(* IEC 61131-3 sources: JingjiangArm/moonboxpro_arm_8.4/Application/Application/任务列表/TensionTask/张力控制/收放料/放料卷径相关/卷径估计, 7 files *)

(* ---- KS_GetFilmThickNessByEstDiaFunc.st ---- *)
(*@CES
Name=KS_GetFilmThickNessByEstDiaFunc
Type=FunctionBlock
TypeGuid=6f9dac99-8de1-4efc-8465-68ac443b7d08
Guid=9700b421-fab0-4030-bfa4-7fb145ef1e2a
HasDeclaration=True
HasImplementation=True
*)
{DECLARATION}
FUNCTION KS_GetFilmThickNessByEstDiaFunc : BOOL
(*2023.12.02.095036 通过估计函数获取料膜厚度@目前主要只应用于接料时的10s不进行卷径补偿部分。
自动获取的方式是
*在开机印刷后超过一定的速度并且处于匀速段
*等待一定的时间后
*持续运行一定的时间后计算这段时间的平均值作为自动的厚度值*)
(*2024.03.16.101611 在停止计算的时候写入初始厚度值|
防止上次料膜太厚计算出的值和本次的薄料厚度差别太大引起异常。厚度值比实际小,对于接料影响会小一些*)
(*2024.7.24.124217 逻辑优化*)
VAR_INPUT
	i_xGetFilmThicknessEn:BOOL;(*自动获取厚度使能@印刷到达一定速度-非调试模式*)
	i_xGetFilmThickNessAuto:BOOL;(*自动获取标志@有效了就通过估计的厚度值获得。无效则通过手动输入获取*)

	i_byWaitTime_Min:BYTE:=1;(*自动满足条件后等待的时间@经过这段时间后开始计算@min*)
	i_byContinuousTime_Min:BYTE:=5;(*持续计算的时间@min*)
	i_byShakeThreshold:BYTE:=10;(*抖动阈值(最值差值法)@丝*)

	i_xEstiThikcknessValid:BOOL;(*估计的厚度值有效*)
	i_rEstiThickness:REAL;(*估计的厚度值@mm*)

	(*2024.03.16.101417*)
	i_rThickness_Init:REAL;(*初始厚度@用于初始化|在退出计算的时候写入该值*)

	i_pxAutoGetDne:POINTER TO BOOL;(*自动获取成功了*)
	i_prThickness:POINTER TO REAL;(*获取的厚度值@mm*)
	i_prTotalThickness:POINTER TO REAL;(*统计的总的厚度值@用于平均处理*)
	i_pudiTotalNum:POINTER TO UDINT;(*统计的次数值@用于平均处理*)
	i_prThickness_Max:POINTER TO REAL;
	i_prThickness_Min:POINTER TO REAL;
	i_ptLastTime:POINTER TO TIME;(*计时使用*)
END_VAR
VAR
	xAutoGetDne: BOOL;
	rThickness: REAL;
	rEstiThickness: REAL;
	rTotalThickness: REAL;
	udiTotalNum: UDINT;
	rThickness_Max: REAL;
	rThickness_Min: REAL;
	rThickness_Manu: REAL;
	tLastTime: TIME;
	tTemp:TIME;
	xEstiThikcknessValid: BOOL;
	rThickness_Init: REAL;(*2024.03.16.101525*)
END_VAR
{IMPLEMENTATION}
(*指针变量写入到临时变量*)
IF i_pxAutoGetDne <>0 THEN
	xAutoGetDne:=i_pxAutoGetDne^;
END_IF
IF i_prThickness<>0 THEN
	rThickness:=i_prThickness^;
END_IF
IF i_prTotalThickness<>0 THEN
	rTotalThickness:=i_prTotalThickness^;
END_IF
IF i_pudiTotalNum<>0 THEN
	udiTotalNum:=i_pudiTotalNum^;
END_IF
IF i_prThickness_Max<>0 THEN
	rThickness_Max:=i_prThickness_Max^;
END_IF
IF i_prThickness_Min<>0 THEN
	rThickness_Min:=i_prThickness_Min^;
END_IF
IF i_ptLastTime<>0 THEN
	tLastTime:=i_ptLastTime^;
END_IF

xEstiThikcknessValid:=i_xEstiThikcknessValid;
rEstiThickness:=i_rEstiThickness;
IF rEstiThickness<=0 OR
	rEstiThickness>=1 THEN(*1MM厚度的几乎没见过，这个只是为了别错的太离谱*)
	xEstiThikcknessValid:=FALSE;(*认为无效|复位所有内容,如果恢复了则重新计算-已经计算完成了就保持吧*)
END_IF

(*2024.03.16.101532*)
rThickness_Init:=i_rThickness_Init;
IF rThickness_Init=0 THEN
	rThickness_Init:=0.02;
END_IF

(*通过估计获取到的厚度值计算*)
(*逻辑处理*)
IF i_xGetFilmThickNessAuto AND(*使用自动获取的方式*)
	xEstiThikcknessValid THEN(*获取估计的厚度值@无效就按照手动输入处理*)
	IF i_xGetFilmThicknessEn AND(*可以自动运算了*)
		NOT xAutoGetDne THEN(*未完成*)
		(*2024.03.16.101150*)
		IF tLastTime=T#0MS THEN(*开始的时候记录时间*)
			tLastTime:=TIME();
		END_IF

		tTemp:=DWORD_TO_TIME(BYTE_TO_DWORD(i_byWaitTime_Min)*60*1000);(*转换为ms*)
		IF TIME()-tLastTime>tTemp THEN(*等待时间够了*)
			tTemp:=DWORD_TO_TIME(BYTE_TO_DWORD(i_byWaitTime_Min+i_byContinuousTime_Min)*60*1000);(*转换为ms*)
			(*累计厚度值*)
			udiTotalNum:=udiTotalNum+1;
			rTotalThickness:=rTotalThickness+rEstiThickness;
			(*记录最大值和最小值*)
			IF rThickness_Max<rEstiThickness THEN
				rThickness_Max:=rEstiThickness;
			END_IF
			IF rThickness_Min>rEstiThickness THEN
				rThickness_Min:=rEstiThickness;
			END_IF

			(*记录的时间到了@检查最大和最小值偏差是否符合要求*)
			IF TIME()-tLastTime>tTemp THEN
				(*符和要求|写入*)
				IF (rThickness_Max-rThickness_Min)<=BYTE_TO_REAL(i_byShakeThreshold)/100.0 THEN
					IF udiTotalNum<>0 THEN
						rThickness:=LREAL_TO_REAL(rTotalThickness/UDINT_TO_LREAL(udiTotalNum));
					ELSE;(*保持之前的值*)
					END_IF
					xAutoGetDne:=TRUE;(*都认为完成了*)
				ELSE(*数据不可靠@重新统计|更新记录的时间信息*)
					tLastTime:=TIME();
				END_IF
			END_IF
		ELSE(*时间还没等够呢|清除无用的变量*)
			udiTotalNum:=0;
			rTotalThickness:=0;
			rThickness_Max:=0;
			rThickness_Min:=999;(*初始化为了较大值*)
		END_IF
	ELSE(*状态还不合适的时候|清除无用的变量*)
		udiTotalNum:=0;
		rTotalThickness:=0;
		rThickness_Max:=0;
		rThickness_Min:=999;(*初始化为了较大值*)
		(*2024.03.16.101249  清零时间@开始的时候会记录*)
(*		tLastTime:=TIME();*)
		(*不再运算的时候复位下*)
		(*2024.7.24.130213 优化*)
		IF NOT i_xGetFilmThicknessEn THEN
			xAutoGetDne:=FALSE;
			IF tLastTime<>T#0MS THEN(*用于标记进入过计算逻辑*)
				tLastTime:=T#0MS;
				rThickness:=rThickness_Init;(*退出运算的时候写入初始厚度值*)
			END_IF
		END_IF
	END_IF
ELSE(*非自动获取的@手动输入*)
	udiTotalNum:=0;
	rTotalThickness:=0;
	rThickness_Max:=0;
	rThickness_Min:=999;(*初始化为了较大值*)
	IF NOT i_xGetFilmThickNessAuto THEN(*不自动获取的时候复位*)
		xAutoGetDne:=FALSE;
		(*2024.7.24.125804|*)
		IF tLastTime<>T#0MS THEN(*用于标记进入过计算逻辑*)
			tLastTime:=T#0MS;
			rThickness:=rThickness_Init;(*退出运算的时候写入初始厚度值*)
		END_IF
	END_IF
END_IF

(*1MM厚度的几乎没见过，这个只是为了别错的太离谱*)
IF rThickness<=0 OR
	rThickness>=1 THEN
	rThickness:=rThickness_Init;
END_IF

(*临时变量写入到指针变量*)
IF i_pxAutoGetDne <>0 THEN
	i_pxAutoGetDne^:=xAutoGetDne;
END_IF
IF i_prThickness<>0 THEN
	i_prThickness^:=rThickness;
END_IF
IF i_prTotalThickness<>0 THEN
	i_prTotalThickness^:=rTotalThickness;
END_IF
IF i_pudiTotalNum<>0 THEN
	i_pudiTotalNum^:=udiTotalNum;
END_IF
IF i_prThickness_Max<>0 THEN
	i_prThickness_Max^:=rThickness_Max;
END_IF
IF i_prThickness_Min<>0 THEN
	i_prThickness_Min^:=rThickness_Min;
END_IF
IF i_ptLastTime<>0 THEN
	i_ptLastTime^:=tLastTime;
END_IF

(* ---- KS_InitEstPara.st ---- *)
(*@CES
Name=KS_InitEstPara
Type=FunctionBlock
TypeGuid=6f9dac99-8de1-4efc-8465-68ac443b7d08
Guid=ee2b4dc0-cfeb-471c-b1f7-6492871368b6
HasDeclaration=True
HasImplementation=True
*)
{DECLARATION}
FUNCTION KS_InitEstPara : BOOL(*初始化估计参数*)
VAR_INPUT
	i_rInitRadius:REAL:=200;(*估计卷半径初始值-mm*)
	i_rInitThickNess:REAL:=0;(*估计厚度初始值*)
	i_parPh:POINTER TO ARRAY [1..3,1..3] OF REAL;(*矩阵地址3X3*)
	i_parXh:POINTER TO ARRAY [1..3] OF REAL;(*矩阵1x3-Xh[1]为估计的卷径(半径-mm),Xh[2]为估计的厚度,Xh[3]为估计的张力 *)
END_VAR
VAR
	(*初始取值*)
	(*估计算法使用了矩阵计算|下面数组实际是矩阵定义*)
	arPh:ARRAY [1..3,1..3] OF REAL:=[1,0,0,0,1,0,0,0,0];
END_VAR
{IMPLEMENTATION}
IF i_parPh<>0 AND
	i_parXh<>0 THEN
	(*进行初始化*)
	i_parPh^:=arPh;
	i_parXh^[1]:=i_rInitRadius;
	i_parXh^[2]:=i_rInitThickNess;
	i_parXh^[3]:=0;
END_IF

(* ---- LowPass.st ---- *)
(*@CES
Name=LowPass
Type=FunctionBlock
TypeGuid=6f9dac99-8de1-4efc-8465-68ac443b7d08
Guid=d3642d54-f54d-4ba9-a90e-82a081cd60e8
HasDeclaration=True
HasImplementation=True
*)
{DECLARATION}
FUNCTION LowPass : BOOL
(*
	功能：一阶低通滤波器   截止频率1rad/s
	输入：计算的补偿量
	输出：滤波后补偿量
*)
VAR_INPUT

	i_rInput:REAL;(*摆臂输出模拟量*)
	i_prOutput: POINTER TO REAL;(*控制器输出转速(r/min)-绝对值*)
	i_parUk:POINTER TO ARRAY [1..2] OF REAL;(*输入寄存器 [U(k);U(k-1)]*)
	i_parYk:POINTER TO ARRAY [1..2] OF REAL;(*输出寄存器[Y(k);Y(k-1)]*)

	(*2023.09.27.222339 增加了截止频率的输入设置*)
	i_rWc:REAL;
	i_iCycleTime_Plc: INT;
END_VAR

VAR
	rTs:REAL :=0.02;

	rAp:REAL :=1.0;  (*%通带允许的最大衰减 dB*)
	rWc:REAL :=2.0;  (*%截止频率rad/s,一般取1，(一般放卷系统的截止频率为1rad/s),若补偿效果差，可以加大，若发散，则减小*)

	rE:REAL :=0;
	rA0:REAL :=0;
	rB0:REAL :=0;
	rA1:REAL :=0;
	rB1:REAL :=0;

	rTemp:REAL :=0;
END_VAR
{IMPLEMENTATION}
(*2023.09.27.222448 增加截止频率的赋值*)
rWc:=i_rWc;
IF rWc<=0 THEN
	rWc:=2;
END_IF
rTs:=INT_TO_REAL(i_iCycleTime_Plc)/1000.0;(*2024.12.3.103753 周期通过变量计算*)
(*参数*)
rTemp :=rAp/10.0;
rTemp :=LREAL_TO_REAL(EXPT(10.0,rTemp));
rE :=SQRT(rTemp-1.0);

rA0:=rWc*rTs;
rA1:=rWc*rTs;

rB0 :=rWc*rTs-2.0*rE;
rB1 :=rWc*rTs+2.0*rE;

(*差分计算*)
i_parUk^[1] :=i_rInput;
i_parYk^[1] :=1/rB1*(rA1*i_parUk^[1]+rA0*i_parUk^[2]-rB0*i_parYk^[2]);

(*更新寄存器*)
i_parUk^[2] :=i_parUk^[1];

i_parYk^[2] :=i_parYk^[1];

(*输出*)
i_prOutput^ :=i_parYk^[1];

(* ---- MatProduct.st ---- *)
(*@CES
Name=MatProduct
Type=FunctionBlock
TypeGuid=6f9dac99-8de1-4efc-8465-68ac443b7d08
Guid=c51cd6fe-fb5a-47c0-a409-be36c7f0e134
HasDeclaration=True
HasImplementation=True
*)
{DECLARATION}
(*需要预先输入：输入矩阵的维数，输出矩阵的维数*)
FUNCTION MatProduct : REAL
VAR_INPUT
	LMat_Row:INT;
	LMat_Col:INT;
	RMat_Row:INT;
	RMat_Col:INT;
	pLMat_Member:POINTER TO  REAL;
	pRMat_Member:POINTER TO  REAL;
	pOutMat_Member:POINTER TO  REAL;
END_VAR
VAR
	iN: INT;
	iJ: INT;
	iK: INT;
	pRMat_temp:POINTER TO  REAL;
	pLMat_temp:POINTER TO  REAL;
	rTwmp1: REAL;
	DW: DWORD;
	rTwmp2: REAL;
	WordLength:DWORD;
END_VAR

{IMPLEMENTATION}
IF pRMat_Member=0 OR pLMat_Member=0 THEN
	RETURN;
END_IF
(*SysMemSet(i_pPh,0,4*9);*)
WordLength:=REAL_TO_DWORD(SIZEOF(pLMat_Member^));
FOR iN:=0 TO LMat_Row-1 BY +1 DO
	FOR iJ:=0 TO RMat_Col-1 BY +1 DO
             pOutMat_Member^:=0;
		FOR iK:=0 TO LMat_Col-1 BY +1 DO
			DW:=INT_TO_DWORD(iN*LMat_Col+iK);
                    pLMat_temp:=pLMat_Member+DW*WordLength;
			rTwmp1:=pLMat_temp^;

			DW:=INT_TO_DWORD(iJ+iK*RMat_Col);
			pRMat_temp:=pRMat_Member+DW*WordLength;
			rTwmp2:=pRMat_temp^;
                   pOutMat_Member^:= pOutMat_Member^+pLMat_temp^*pRMat_temp^;
		END_FOR
		pOutMat_Member:=pOutMat_Member+WordLength;
	END_FOR
END_FOR
(*pOutMat_Member:=pOutMat_Member-WordLength*(LMat_Row*RMat_Col-1);*)

(* ---- RadiEst.st ---- *)
(*@CES
Name=RadiEst
Type=FunctionBlock
TypeGuid=6f9dac99-8de1-4efc-8465-68ac443b7d08
Guid=78b04f11-b967-4930-a408-d7c5f7f7845f
HasDeclaration=True
HasImplementation=True
*)
{DECLARATION}
FUNCTION RadiEst : REAL
VAR_INPUT
	i_xFilmToBig:BOOL;(*TRUE:料膜变大；FALSE:料膜变小*)
	i_Wu:REAL;(*放料转速(RPM)*)
	i_Vt:REAL;(*牵引线速度,(mm/s)*)
	i_Tf:REAL;(*张力摆臂反馈(V)*)
	i_EaL:REAL;(*i_EaL=10.08，弹性模量(N/m^2)*横截面积(m^2)/料长(mm)*)
	i_Ts:REAL;(*采样周期(s)*)
	i_Para_Tf:REAL;(*张力迭代参数|1*)
	i_Para_R:REAL;(*卷径迭代参数|100*)
	i_pPh:POINTER TO  REAL;(*二维数组Ph指针*)
	i_pXh:POINTER TO  REAL;(*上一个周期估计状态向量Xh指针*)
END_VAR
VAR
	pPtemp3_1:POINTER TO  REAL;(*一维数组临时指针*)
	pPtemp3_3a:POINTER TO  REAL;(*二维数组P和Ph的临时指针*)
	pPtemp3_3b:POINTER TO  REAL;(*二维数组P和Ph的临时指针*)
	pXtemp:POINTER TO REAL;
	pAp:POINTER TO  REAL;(*二维数组A指针*)
	pCp:POINTER TO  REAL;(*二维数组A指针*)
	pApt: POINTER TO REAL;
	pK:POINTER TO REAL;
	pX:POINTER TO REAL;(*状态向量指针*)
	pP:POINTER TO REAL;
	pTemp:POINTER TO REAL;
	Apt:ARRAY [1..3,1..3] OF REAL:=[0,0,0,0,0,0,0,0,0];
	Ap:ARRAY [1..3,1..3] OF REAL:=[0,0,0,0,0,0,0,0,0];
	Cp:ARRAY [1..3] OF REAL:=[0,0,1];
	P:ARRAY [1..3,1..3] OF REAL;(*:=0,0,0,0,0,0,0,0*)
	Ptemp3_3a:ARRAY [1..3,1..3] OF REAL;(*:=0,0,0,0,0,0,0,0*)
	Ptemp3_3b:ARRAY [1..3,1..3] OF REAL;(*:=0,0,0,0,0,0,0,0*)
	Ptemp3_1:ARRAY [1..3] OF REAL;(*:=0,0,0,0,0,0,0,0*)
	K:ARRAY [1..3] OF REAL:=[0,0,0];
	X:ARRAY [1..3] OF REAL:=[0,0,0];
	Xtemp:ARRAY [1..3] OF REAL:=[0,0,0];
	iN:INT;
	Temp:REAL;

	parTemp:POINTER TO ARRAY [1..3,1..3] OF REAL;
	iCoeff: INT;
END_VAR
{IMPLEMENTATION}
(*将函数中的数组和指针关联*)
pAp:=ADR(Ap);
pApt:=ADR(Apt);
pCp:=ADR(Cp);
pPtemp3_1:=ADR(Ptemp3_1);
pPtemp3_3a:=ADR(Ptemp3_3a);
pPtemp3_3b:=ADR(Ptemp3_3b);
pK:=ADR(K);
pXtemp:=ADR(Xtemp);
pP:=ADR(P);
pX:=ADR(X);
(*针对卷径变化方向增加|标志切换*)
IF i_xFilmToBig THEN(*卷径变大了*)
	iCoeff:=1;
ELSE(*卷径变小了*)
	iCoeff:=-1;
END_IF

(*给Ap,Apt,Cp,X赋值*)
Ap[1,1]:=1 ; Ap[1,2]:=iCoeff*i_Wu*i_Ts/60 ; Ap[2,2]:=1 ; Ap[3,1]:=LREAL_TO_REAL(iCoeff*i_EaL*i_Ts*i_Wu/60*2*gc_lrPi) ; Ap[3,3]:=1;
Apt[1,1]:=1 ; Apt[2,1]:=iCoeff*i_Wu*i_Ts/60 ; Apt[2,2]:=1 ; Apt[1,3]:=LREAL_TO_REAL(iCoeff*i_EaL*i_Ts*i_Wu/60*2*gc_lrPi) ; Apt[3,3]:=1;
Cp[3]:=1;
(*Ph=APA'+Q*)
MatProduct(3,3,3,3,pAp,i_pPh,pPtemp3_3a);
MatProduct(3,3,3,3,pPtemp3_3a,pApt,i_pPh);
pTemp:=i_pPh+REAL_TO_DWORD(8*4);
pTemp^:=pTemp^+i_Para_Tf;
(*K=Ph*C'/(R+C*Ph*C')*)
MatProduct(3,3,3,1,i_pPh,pCp,pK);
pTemp:=i_pPh+REAL_TO_DWORD(8*4);
Temp:=i_Para_R+pTemp^;
FOR iN:=1 TO 3 BY +1 DO
K[iN]:=K[iN]/Temp;
END_FOR
(*X=Ax+Bu*)
MatProduct(3,3,3,1,pAp,i_pXh,pXtemp);
Xtemp[3]:=Xtemp[3]+i_Ts*i_EaL*i_Vt*(-iCoeff);
X:=Xtemp;
(*Xh=X+K(y-CX)*)
Temp:=0;
Temp:=i_Tf-X[3];
FOR iN:=1 TO 3 BY +1 DO
pTemp:=i_pXh+INT_TO_DWORD(4*(iN-1));
pTemp^:=X[iN]+Temp*K[iN];
END_FOR
(*P=(I-KC)Ph*)
Cp[3]:=-1;
MatProduct(3,1,1,3,pK,pCp,pPtemp3_3a);
Ptemp3_3a[1,1]:=1.0+Ptemp3_3a[1,1];
Ptemp3_3a[2,2]:=1.0+Ptemp3_3a[2,2];
Ptemp3_3a[3,3]:=1.0+Ptemp3_3a[3,3];
pPtemp3_3b:=i_pPh;
(*MatProduct(3,3,3,3,pPtemp3_3a,pPtemp3_3b,i_pPh);将估计协方差矩阵传出*)
MatProduct(3,3,3,3,pPtemp3_3a,i_pPh,pP);(*将估计协方差矩阵传出*)
(*g_Ph:=P;*)
parTemp:=i_pPh;
parTemp^:=P;

(* ---- KS_FB_CalcDiamOfFilmVol.st ---- *)
(*@CES
Name=KS_FB_CalcDiamOfFilmVol
Type=FunctionBlock
TypeGuid=6f9dac99-8de1-4efc-8465-68ac443b7d08
Guid=aa4e7948-893a-473e-86a9-5c9051eef5bc
HasDeclaration=True
HasImplementation=True
*)
{DECLARATION}
FUNCTION_BLOCK KS_FB_CalcDiamOfFilmVol(*卷径计算*)
VAR_INPUT
	i_xEnable: BOOL;
	i_lrFilmVelocity:LREAL;(*料膜速度*)
	i_lrUnWind_Velocity:LREAL;(*放料速度参数*)
	i_lrWind_Velocity :LREAL;(*收料速度参数*)
	i_lrAlarm_Diameter: LREAL ;(*报警卷径*)
	i_xUnWind_CutFinished: BOOL;(*放料裁切完成*)
	i_xWind_CutFinished: BOOL;(*收料裁切完成*)
	i_CycleTime:INT;(*程序循环时间*)
	i_xRollerPress_Uw:BOOL;(*全体合压标志*)
	i_xMachineRev:BOOL;(*整机反转标志*)
	(*2021.8.26.173437 增加了预估卷径以后添加的参数*)
	i_rDiaAcT_Uw:REAL;(*放料实际当前卷径*)
	i_rDiaAcT_Rw:REAL;(*放料实际当前卷径*)
END_VAR
VAR_OUTPUT
	o_xEno: BOOL;
	o_iErNo: INT;
	o_xFlag_AlarmDiameter: BOOL;
END_VAR
VAR_IN_OUT
	rUnWind_Diameter:REAL;(*放料卷径*)
	rWind_Diameter:REAL;(*收料卷径*)
END_VAR
VAR
	temp1: LREAL;
	temp2: LREAL;
(*2016年5月26日 14:45:08*)
	rUnWind_DiameterArr: ARRAY [1..200] OF LREAL;		(*放料计算卷径*)
	rWind_DiameterArr: ARRAY [1..200] OF LREAL;		(*收料计算卷径*)
	iNum: INT := 150;(*卷径平均次数*)
	lrUnWind_Velocity: ARRAY[1..200] OF LREAL;
	lrWind_Velocity: ARRAY[1..200] OF LREAL;
	iEven_Num: INT := 5;(*速度平均次数*)
	lrSum_UnWind_Velocity: LREAL;
	lrSum_Wind_Velocity: LREAL;	(*  *)
	lrSum_UnWind_Diameter: LREAL;
	lrSum_Wind_Diameter: LREAL;
	iN: INT;
	Init: BOOL;(*收放料速度、卷径数组初始化标志*)
	lrUnWind_Dia: LREAL;(*放料平均卷径*)
	lrWind_Dia: LREAL;(*收料平均卷径*)

	iCalDiameter: INT:=20;(*卷径计算间隔时间ms*)
	iCalDiameterCycleCount:INT:=1;(*卷径计算周期计数*)

	iUnwindDia_Min:INT:=80;(*放料最小卷径*)
	iUnwindDia_Max:INT:=1600;(*放料最大卷径*)
	iwindDia_Min:INT:=80;(*收料最小卷径*)
	iwindDia_Max:INT:=1600;(*收料最大卷径*)

	iTemp: INT;(*控制卷径计算方向的*)
	uiUpdateDia: UINT;
	uiCount: UINT;(*计数，用来确定卷径变化已经稳定，防止卷径报警异常输出*)
	lrStep_Uw: LREAL;
	lrTime_Temp: LREAL := 5000;
	lrStep_Rw: LREAL;
END_VAR

{IMPLEMENTATION}
o_xEno:= i_xEnable;
o_iErNo:= 0;

(*需要放在fb_Vel_TO_Vol功能块后，因为在fb_Vel_TO_Vol功能块中进行卷径的切换。*
*	同时要放在收放料裁切换料标志清零之前                                   *)
IF i_xEnable THEN
	IF i_xUnWind_CutFinished OR  i_xWind_CutFinished THEN(*放料或者收料裁切完成，置Init标志为false*)
		Init:=FALSE;
	END_IF
(*2020.9.30.094859|liu.yt删除该处赋值变量|
	iEven_Num:=150;
*)
	IF iCalDiameterCycleCount >=iCalDiameter/i_CycleTime THEN(*卷径计算周期条件*)
		iCalDiameterCycleCount:=1;
		IF NOT Init THEN(*收放料速度、卷径数组初始化*)
			Init:=TRUE;
			FOR iN:=1 TO iEven_Num BY 1 DO
				lrUnWind_Velocity[iN]:=i_lrUnWind_Velocity;
				lrWind_Velocity[iN]:=i_lrWind_Velocity;
			END_FOR
			FOR iN:=1 TO iNum BY 1 DO
				rUnWind_DiameterArr[iN]:=rUnWind_Diameter;
				rWind_DiameterArr[iN]:=rWind_Diameter;
			END_FOR
			temp1:=i_lrFilmVelocity;
			temp2:=i_lrFilmVelocity;
		END_IF

	(*计算平均线速度*)
		FOR iN:=iEven_Num TO 2 BY -1 DO
			lrUnWind_Velocity[iN] := lrUnWind_Velocity[iN-1];
			lrWind_Velocity[iN] := lrWind_Velocity[iN-1];
		END_FOR
		lrUnWind_Velocity[1]:=i_lrUnWind_Velocity;
		lrWind_Velocity[1]:=i_lrWind_Velocity;
		lrSum_UnWind_Velocity := 0;
		lrSum_Wind_Velocity := 0;
		FOR iN:=1 TO iEven_Num BY 1 DO
			lrSum_UnWind_Velocity:=lrSum_UnWind_Velocity+lrUnWind_Velocity[iN];
			lrSum_Wind_Velocity:=lrSum_Wind_Velocity+lrWind_Velocity[iN];
		END_FOR
		temp1 := lrSum_UnWind_Velocity / iEven_Num;(*计算放料平均速度*)
		temp2 := lrSum_Wind_Velocity / iEven_Num;(*计算收料平均速度*)
	(*计算平均卷径*)
		FOR iN:=iNum TO 2 BY -1 DO
			rUnWind_DiameterArr[iN] := rUnWind_DiameterArr[iN-1];
			rWind_DiameterArr[iN] := rWind_DiameterArr[iN-1];
		END_FOR

(*计算收放料直径用于计算料膜平均直径*)

		IF temp1<>0 THEN(*卷径=料膜速度/角速度*)
			rUnWind_DiameterArr[1]:=i_lrFilmVelocity/temp1/3.14159*1000;
		END_IF

		IF rUnWind_DiameterArr[1] <iUnwindDia_Min THEN
			rUnWind_DiameterArr[1]:=iUnwindDia_Min;
		END_IF

		IF rUnWind_DiameterArr[1] >iUnwindDia_Max THEN
			rUnWind_DiameterArr[1]:=iUnwindDia_Max;
		END_IF

		IF temp2<>0 THEN	(*卷径=料膜速度/角速度*)
			rWind_DiameterArr[1]:=i_lrFilmVelocity/temp2/3.14159*1000;
		END_IF

		IF rWind_DiameterArr[1] <iwindDia_Min THEN
			rWind_DiameterArr[1]:=iwindDia_Min;
		END_IF

		IF rWind_DiameterArr[1] >iwindDia_Max THEN
			rWind_DiameterArr[1]:=iwindDia_Max;
		END_IF

		lrSum_UnWind_Diameter := 0;
		lrSum_Wind_Diameter := 0;
		FOR iN:=1 TO iNum BY 1 DO
			lrSum_UnWind_Diameter := lrSum_UnWind_Diameter + rUnWind_DiameterArr[iN];
			lrSum_Wind_Diameter := lrSum_Wind_Diameter + rWind_DiameterArr[iN];
		END_FOR
		lrUnWind_Dia:=lrSum_UnWind_Diameter/iNum;(*计算放料平均卷径值*)
		lrWind_Dia:=lrSum_Wind_Diameter/iNum;(*计算收料平均卷径值*)

(*整机反转时候卷径计算控制*)
		IF i_xMachineRev THEN
			iTemp:=-1;
		ELSE
			iTemp:=1;
		END_IF

		IF i_lrFilmVelocity>=10 THEN(*角速度控制算法的时候开机就计算卷径，线速度算法需要大于15M/MIN时候计算*)
			uiUpdateDia:=uiUpdateDia+1;(*卷径更新计数*)
			IF uiUpdateDia>=10 THEN(*200更新一次*)
				IF NOT i_xRollerPress_Uw THEN (*放料胶辊未合压了*)
					(*防止由于裁切换料的时候 可能会导致卷径计算不准确，进行卷径切换的时候会出错，所以在此时不再计算保持之前的值*)
					IF lrTime_Temp<>0 THEN
						lrStep_Uw:= ABS(rUnWind_Diameter-lrUnWind_Dia)*i_CycleTime*uiUpdateDia/lrTime_Temp;
						IF lrStep_Uw<(*0.1 *)0.2 THEN(*|从数据中发现为0.1时不能跟上卷径的变化*)
							lrStep_Uw:=(*0.1*)0.2;
						ELSE;
						END_IF
					END_IF
					IF ABS( rUnWind_Diameter-lrUnWind_Dia)<=50 THEN
						IF iTemp*(rUnWind_Diameter - lrUnWind_Dia) > lrStep_Uw THEN
							rUnWind_Diameter := rUnWind_Diameter  - lrStep_Uw*iTemp;
						ELSIF  -iTemp*(rUnWind_Diameter - lrUnWind_Dia) >lrStep_Uw THEN
							rUnWind_Diameter := rUnWind_Diameter  + lrStep_Uw*iTemp;
						ELSE
							rUnWind_Diameter:=lrUnWind_Dia;
						END_IF
					ELSE
						rUnWind_Diameter:=lrUnWind_Dia;
					END_IF
				END_IF

				IF lrTime_Temp<>0 THEN
					lrStep_Rw:= ABS(rWind_Diameter-lrWind_Dia)*20*uiUpdateDia/lrTime_Temp;
					IF lrStep_Rw<(*0.1*)0.2 THEN(*1S-0.5mm*)(*将卷径最小变化率改为0.3即1.5mm/s.|从数据中发现为0.1时不能跟上卷径的变化*)
						lrStep_Rw:=(*0.1*)0.2;
					ELSE;
					END_IF
				END_IF
				IF ABS( rWind_Diameter-lrWind_Dia)<=50 THEN
					IF iTemp*(rWind_Diameter - lrWind_Dia) > lrStep_Rw THEN
						rWind_Diameter := rWind_Diameter  - lrStep_Rw*iTemp;
					ELSIF  -iTemp*(rWind_Diameter - lrWind_Dia) > lrStep_Rw THEN
						rWind_Diameter := rWind_Diameter  + lrStep_Rw*iTemp;
					ELSE
						rWind_Diameter:=lrWind_Dia;
					END_IF
				ELSE
					rWind_Diameter:=lrWind_Dia;
				END_IF
				uiUpdateDia:=0;
			END_IF

(*卷径报警输出*)
			IF NOT i_xMachineRev THEN(*整机正转时候*)
				IF  i_rDiaAcT_Uw <= i_lrAlarm_Diameter+2 THEN(*+2是为了防止放料计算的卷径抖动，重复触发报警*)
					IF i_rDiaAcT_Uw <= i_lrAlarm_Diameter THEN
						IF uiCount>=250 THEN(*连续5S放料卷径都小于报警卷径则认为需要报警*)
							o_xFlag_AlarmDiameter := TRUE;
						ELSE
							uiCount:=uiCount+1;
						END_IF
					ELSE
						uiCount:=0;
					END_IF
				ELSE
					uiCount:=0;
					o_xFlag_AlarmDiameter := FALSE;
				END_IF
			END_IF

			IF  i_xMachineRev THEN(*整机反转时候*)
				IF  i_rDiaAcT_Rw <= i_lrAlarm_Diameter+2 THEN(*+2是为了防止放料计算的卷径抖动，重复触发报警*)
					IF i_rDiaAcT_Rw <= i_lrAlarm_Diameter THEN
						IF uiCount>=250 THEN(*连续5S放料卷径都小于报警卷径则认为需要报警*)
							o_xFlag_AlarmDiameter := TRUE;
						ELSE
							uiCount:=uiCount+1;
						END_IF
					ELSE
						uiCount:=0;
					END_IF
				ELSE
					uiCount:=0;
					o_xFlag_AlarmDiameter := FALSE;
				END_IF
			END_IF

		END_IF

		IF rUnWind_Diameter <= iUnwindDia_Min THEN
			rUnWind_Diameter := iUnwindDia_Min;
		END_IF
		IF rUnWind_Diameter >= iUnwindDia_Max THEN
			rUnWind_Diameter := iUnwindDia_Max;
		END_IF

		IF rWind_Diameter <= iwindDia_Min THEN
			rWind_Diameter := iwindDia_Min;
		END_IF
		IF rWind_Diameter >= iwindDia_Max THEN
			rWind_Diameter := iwindDia_Max;
		END_IF
	ELSE
		iCalDiameterCycleCount:=iCalDiameterCycleCount+1;
	END_IF
ELSE
	o_xFlag_AlarmDiameter := FALSE;
	Init:=FALSE;
	iCalDiameterCycleCount:=1;
	uiUpdateDia:=0;(*卷径更新周期计数*)
	uiCount:=0;
END_IF

(* ---- KS_FB_EstimationByVel.st ---- *)
(*@CES
Name=KS_FB_EstimationByVel
Type=FunctionBlock
TypeGuid=6f9dac99-8de1-4efc-8465-68ac443b7d08
Guid=7013804d-3856-4a07-9c38-8f3020ce9a4d
HasDeclaration=True
HasImplementation=True
*)
{DECLARATION}
FUNCTION_BLOCK KS_FB_EstimationByVel(*收放料通过牵引速度(也可以使用料膜速度)以及自己转速估计卷半径以及料膜厚度算法-By.CHEN*)
(*预估之前会重新初始化预估卷径值*)
(*2023.06.08.162623 限制最大卷径增加接口
初始卷径值获取方式可配置*)
(*2023.6.24.101658 重新调整初始卷径的赋值方式@Liu.yt*)
(*2024.01.02.111942优化接口*)
VAR_INPUT
	i_xEn:BOOL;(*估计使能|*)
	i_xFilmToBig:BOOL;(*TRUE:料膜变大；FALSE:料膜变小*)
	i_rFeedBack:REAL;(*摆臂位置反馈位置-V*)
	i_rVel_rpm:REAL;(*估计所需要的当前转速|r/min*)
	i_rVel_mpm:REAL;(*估计所需要的当前速度变量|-线速度m/min*)
	i_xCutDne:BOOL;(*裁切完成标志|只有效一个周期*)
	i_rNewDia:REAL;(*新卷卷直径-mm*)
	i_uiMaxDia:UINT;(*机械最大卷直径-mm*)
	i_uiInitDiam:UINT;(*初始卷直径|=0自动方式设置-mm*)
	i_xTypeGetInitDiam:BOOL;(*方式切换|FALSE=使用停机之前的值|=TRUE 使用固定值*)
	i_rInitThickNess:REAL:=0;(*估计厚度初始值@2023.12.15.234758*)
	i_rInitThickNess_Cut:REAL:=0;(*接料时候估计厚度初始值-接料时候使用之前记录的值@2023.12.15.234758*)
	i_rPara_R:REAL;(*卷径迭代参数|100@2023.12.16.101753*)
	i_iCycleTime_Plc: INT;
END_VAR
VAR_OUTPUT
	o_xEn:BOOL;
	o_rEstThickness:REAL;(*估计的厚度|mm*)
END_VAR
VAR_IN_OUT
	io_rEstDia:REAL;(*估计的卷径-直径mm*)
END_VAR
VAR
	xInitParaDne:BOOL:=FALSE;(*初始化参数完成*)
	(*估计算法使用了矩阵计算|下面数组实际是矩阵定义*)
	arPh:ARRAY [1..3,1..3] OF REAL:=[1,0,0,0,1,0,0,0,0];
	arXh:ARRAY [1..3] OF REAL:=[200,0,0];(*Xh[1]为估计的卷半径,Xh[2]为估计的厚度,Xh[3]为估计的张力*)
	rInitDiam: REAL;(*2023.6.24.101953 初始卷径*)
	uiDiam_Min:UINT:=80;(*最小卷径*)
	rLastInitDiam:REAL;(*初始卷径备份值@发生变化了就更新下*)
	xLastTypeGetInitDiam: BOOL;(*卷径更新方式切换了|更新下*)
END_VAR
{IMPLEMENTATION}
IF i_uiMaxDia < 500 THEN
	i_uiMaxDia:=500;
END_IF

IF i_rPara_R<=0 THEN
	i_rPara_R:=100;
END_IF

IF i_uiInitDiam=0 THEN
	rInitDiam:=(UINT_TO_REAL(i_uiMaxDia)-200)/2.0+200;
ELSE
	rInitDiam:=UINT_TO_REAL(i_uiInitDiam);
END_IF
(*初始值的限值处理*)
IF rInitDiam<uiDiam_Min THEN
	rInitDiam:=uiDiam_Min;
ELSIF rInitDiam>i_uiMaxDia THEN
	rInitDiam:=UINT_TO_REAL(i_uiMaxDia);
END_IF

(*裁切完成了需要更新卷径估计值*)
IF i_xCutDne THEN
	KS_InitEstPara(i_rNewDia/2, i_rInitThickNess_Cut, ADR(arPh), ADR(arXh));(*以新卷半径为基础估计*)
	io_rEstDia:=arXh[1]*2;(*输出为直径*)
END_IF
IF i_xEn THEN(*可以进行估计了|在接换料的时候需要初始化估计参数*)
	(*执行估计算法*)
	RadiEst(
		i_xFilmToBig,
		i_rVel_rpm(*i_Wu*),
		i_rVel_mpm*1000/60(*i_Vt*),
		i_rFeedBack(*i_Tf*),
		1000(*i_EaL*),
		INT_TO_REAL(i_iCycleTime_Plc)/1000(*i_Ts*),
		1(*i_Para_Tf*),
		i_rPara_R(*100*)(*i_Para_R*),(*2023.12.16.101934 修改为了参数*)
		ADR(arPh)(*i_pPh*),
		ADR(arXh)(*i_pXh*));
	io_rEstDia:=arXh[1]*2;(*输出为直径*)
	xInitParaDne:=FALSE;
ELSE(*不使能的时候初始化估计数组*)

	IF rInitDiam<>rLastInitDiam THEN(*初始值发生了变化@重新赋值*)
		xInitParaDne:=FALSE;
	END_IF
	rLastInitDiam:=rInitDiam;(*放到这里应该问题不大。不用在if中再放一次*)

	IF i_xTypeGetInitDiam<>xLastTypeGetInitDiam THEN
		xInitParaDne:=FALSE;
	END_IF
	xLastTypeGetInitDiam:=i_xTypeGetInitDiam;(*放到这里应该问题不大。不用在if中再放一次*)

	IF NOT xInitParaDne THEN
		xInitParaDne:=TRUE;
		(*新方法|2023.06.08.161459*)
		IF i_xTypeGetInitDiam THEN
			KS_InitEstPara(rInitDiam/2, i_rInitThickNess, ADR(arPh), ADR(arXh));(*以新卷半径为基础估计*)
		ELSE
			KS_InitEstPara(io_rEstDia/2, i_rInitThickNess, ADR(arPh), ADR(arXh));(*2022.7.25.165959 初始值修改为之前的值*)
		END_IF
(*		KS_InitEstPara(150, 0, ADR(arPh), ADR(arXh));*)
(*		KS_InitEstPara(200, 0, ADR(arPh), ADR(arXh));*)(* 2021.12.20.100929预估值改为300*)
		io_rEstDia:=arXh[1]*2;(*输出为直径*)
	END_IF
END_IF
(*输出估计的卷半径为直径
以及厚度值*)
o_rEstThickness:=arXh[2];

IF io_rEstDia>=i_uiMaxDia THEN(*输出的估计值进行限值*)
	io_rEstDia:=UINT_TO_REAL(i_uiMaxDia);
ELSIF io_rEstDia<uiDiam_Min THEN
	io_rEstDia:=uiDiam_Min;
END_IF
